(* IEC 61131-3 sources: PortalRobot/Portal_robot/Device/application/ST/ST_CELL, 17 files *)

(* ---- E_CELL_MANAGER_STATE.st ---- *)
{attribute 'qualified_only'}
{attribute 'strict'}
TYPE E_CELL_MANAGER_STATE :
(
	IDLE,
	PLAN_TARGET,
	MAGAZINE_EXECUTE,
	RELEASE_MAGAZINE,
	ROUTE_TO_TARGET,
	RELEASE_ROBOT_COMMAND,
	WAIT_TARGET,
	SERVICE_TARGET,
	SELECT_FALLBACK,
	WAIT_MAGAZINE,
	ERROR,
	MACHINE_FAULT_STOP,
	PRESTART_IDENTIFY,
	WAIT_GRIPPER1_CONTENT,
	WAIT_GRIPPER1_TYPE,
	WAIT_GRIPPER2_CONTENT,
	WAIT_GRIPPER2_TYPE,
	WAIT_START_MACHINE,
	TEST_ABORT_STOP,
	GEOMETRY_WAIT_FREE,
	GEOMETRY_DELIVER,
	GEOMETRY_RELEASE_COMMAND
);
END_TYPE

(* ---- E_CELL_STATE.st ---- *)
{attribute 'qualified_only'}
{attribute 'strict'}
TYPE E_CELL_STATE :
(
	IDLE,
	ROUTE_PAYLOAD,
	SELECT_MACHINE,
	MOVE_TO_MACHINE,
	RELEASE_ROBOT_COMMAND,
	WAIT_MACHINE,
	SERVICE_MACHINE,
	MAGAZINE,
	RELEASE_MAGAZINE,
	WAIT_MAGAZINE,
	ERROR,
	GEOMETRY_WAIT,
	GEOMETRY_TRANSFER
);
END_TYPE

(* ---- ST_BUTTON_STATION_IO_STATUS.st ---- *)
TYPE ST_BUTTON_STATION_IO_STATUS :
STRUCT
	xEmergencyStopPressed : BOOL; // Нормализованный вход: TRUE — грибок нажат
	xButtonPressed        : BOOL; // Нормализованный вход кнопки открытия замка
	xButtonLightOn        : BOOL; // Фактический выход подсветки кнопки
END_STRUCT
END_TYPE

(* ---- ST_CELL_COMMAND.st ---- *)
TYPE ST_CELL_COMMAND :
STRUCT
	stRobot          : ST_ROBOT_COMMAND; // Команда роботу от менеджера ячейки
	uiBlankPayloadType  : UINT; // Тип заготовки в первом захвате
	uiDetailPayloadType : UINT; // Тип готовой детали во втором захвате
	stMagazine       : ST_MAGAZINE_COMMAND; // Команда магазину
	axMachineExecute : ARRAY [1..3] OF BOOL; // Запуск обслуживания выбранного станка
END_STRUCT
END_TYPE

(* ---- ST_CELL_CYCLE_STATUS.st ---- *)
TYPE ST_CELL_CYCLE_STATUS :
STRUCT
	eState              : E_CELL_MANAGER_STATE; // Состояние универсального автомата ячейки
	uiSelectedMachine   : UINT; // Зафиксированный целевой станок
	uiSelectedType      : UINT; // Тип заготовки текущего маршрута
	uiBlankPayloadType  : UINT; // Тип заготовки в первом захвате
	uiDetailPayloadType : UINT; // Тип готовой детали во втором захвате
	iTakeSlot           : SINT; // Зарезервированный слот взятия
	iPutSlot            : SINT; // Зарезервированный слот укладки
	xReturningBlank     : BOOL; // Выполняется возврат заготовки
	axMachineStartPending: ARRAY [1..3] OF BOOL; // Запуск нового цикла ещё подтверждается станком
	auiBlankCount       : ARRAY [1..3] OF UINT; // Заготовки по типам
	auiDetailCount      : ARRAY [1..3] OF UINT; // Готовые детали по типам
	auiFreeCount        : ARRAY [1..3] OF UINT; // Свободные слоты по типам
END_STRUCT
END_TYPE

(* ---- ST_CELL_DIAG.st ---- *)
TYPE ST_CELL_DIAG :
STRUCT
	eState : E_CELL_STATE; // Текущее состояние автомата ячейки
	stWarning : ST_WARNING_EVENT; // Последнее предупреждение менеджера ячейки
END_STRUCT
END_TYPE

(* ---- ST_CELL_ERROR.st ---- *)
TYPE ST_CELL_ERROR :
STRUCT
	BOTH_GRIPPERS_OCCUPIED : BOOL; // Совместимый бит: диагностическая ошибка согласованности захватов
	ROBOT_ERROR            : BOOL; // Ошибка робота во время автоматического цикла
	MAGAZINE_ERROR         : BOOL; // Ошибка магазина во время операции
	MACHINE_ERROR          : BOOL; // Ошибка станка во время обслуживания
	GLOBAL_STOP            : BOOL; // Получена глобальная ошибка ячейки
END_STRUCT
END_TYPE

(* ---- ST_CELL_ERRORS.st ---- *)
TYPE ST_CELL_ERRORS :
STRUCT
	dwErrorActive : DWORD; // Битовая маска активных ошибок
	dwErrorLast   : DWORD; // Битовая маска последних ошибок
	dwAlarmActive : DWORD; // Собственные аварии менеджера ячейки для общего журнала
	stErrorActive : ST_CELL_ERROR; // Расшифровка активных ошибок
	stErrorLast   : ST_CELL_ERROR; // Расшифровка последних ошибок
END_STRUCT
END_TYPE

(* ---- ST_CELL_FAULT_REQUEST.st ---- *)
TYPE ST_CELL_FAULT_REQUEST :
STRUCT
	xEnabled      : BOOL; // Глобальное разрешение диагностической инъекции
	xBothGrippers : BOOL; // Совместимый диагностический импульс ошибки согласованности захватов
END_STRUCT
END_TYPE

(* ---- ST_CELL_SAFETY_DIAG.st ---- *)
TYPE ST_CELL_SAFETY_DIAG :
STRUCT
	stWarning : ST_WARNING_EVENT; // Отклонённые попытки открытия и сброса реле
END_STRUCT
END_TYPE

(* ---- ST_CELL_SAFETY_ERRORS.st ---- *)
TYPE ST_CELL_SAFETY_ERRORS :
STRUCT
	dwErrorActive : DWORD; // Текущие отдельные Safety-причины
	dwErrorLast   : DWORD; // Последняя ненулевая маска для диагностики
	dwAlarmActive : DWORD; // Собственные аварии источника для общего журнала
END_STRUCT
END_TYPE

(* ---- ST_CELL_SAFETY_FAULT_REQUEST.st ---- *)
TYPE ST_CELL_SAFETY_FAULT_REQUEST :
STRUCT
	xEnabled : BOOL; // Общее разрешение диагностических инъекций
	axEmergencyStopStation : ARRAY [1..4] OF BOOL;
	axEmergencyStopCabinet : ARRAY [1..2] OF BOOL;
	xEmergencyStopMpg      : BOOL;
	xPhaseRelayFault       : BOOL;
	xPressureRelayFault    : BOOL;
	xSafetyRelayFault      : BOOL;
	axDoorUnlocked         : ARRAY [1..4] OF BOOL;
END_STRUCT
END_TYPE

(* ---- ST_CELL_SAFETY_STATUS.st ---- *)
TYPE ST_CELL_SAFETY_STATUS :
STRUCT
	xReady                   : BOOL; // Все текущие условия безопасности выполнены
	xGlobalError             : BOOL; // Хотя бы одна текущая Safety-причина активна
	xPhaseRelayOk            : BOOL; // Реле контроля фаз в норме
	xPressureRelayOk         : BOOL; // Реле контроля давления в норме
	xSafetyRelayOk           : BOOL; // Реле безопасности взведено
	xSafetyRelayResetAllowed : BOOL; // Разрешён отдельный импульс сброса реле
	xSafetyRelayResetActive  : BOOL; // Полный секундный импульс сброса реле сейчас активен
	axEmergencyStopReleased  : ARRAY [1..7] OF BOOL; // 4 поста, 2 шкафа, MPG
	axDoorReady              : ARRAY [1..4] OF BOOL; // Замок закрыт либо связанный магазин выключен
	axButtonStationPressed   : ARRAY [1..4] OF BOOL; // Фактический вход кнопки поста, с учётом симуляции
	axButtonStationLightOn   : ARRAY [1..4] OF BOOL; // Выход подсветки кнопки поста
END_STRUCT
END_TYPE

(* ---- ST_CELL_STATUS.st ---- *)
TYPE ST_CELL_STATUS :
STRUCT
	xMagazineExchangeAllowed : BOOL; // Планировщик не держит незавершённый маршрут
	xRunning           : BOOL; // Автоматический цикл запущен
	xStopPending       : BOOL; // Запрошена остановка после безопасного шага
	xBusy              : BOOL; // Менеджер выполняет автоматический цикл
	xWaitingMachine    : BOOL; // Ожидание доступного станка
	xWaitingMagazine   : BOOL; // Ожидание пополнения или освобождения магазина
	xError             : BOOL; // Менеджер ячейки находится в ошибке
	xReadyToStart      : BOOL; // Выполнены все условия запуска автоматического цикла
	xStartAllowed      : BOOL; // Кнопка запуска или отмены ожидающей остановки доступна
	xStopAllowed       : BOOL; // Кнопка остановки автоматического цикла доступна
	xResetAllowed      : BOOL; // Кнопка общего сброса доступна
	xManualAllowed     : BOOL; // Кнопка перехода в ручной режим доступна
	xAutomaticAllowed  : BOOL; // Кнопка перехода в автоматический режим доступна
	xDrivesReady       : BOOL; // Приводы и группа осей готовы к движению
	xRobotReady        : BOOL; // Робот готов принять команду
	xMagazineReady     : BOOL; // Магазин готов к работе с роботом
	xSafetyHomeRequired: BOOL; // Повторный запуск разрешён только из HOME_SAFETY
	xRobotAtSafetyHome : BOOL; // Фактические координаты находятся в диапазоне HOME_SAFETY
	xStartCheckCellIdle          : BOOL; // Менеджер ячейки готов принять новый запуск
	xStartCheckAutomaticMode     : BOOL; // Выбран автоматический режим
	xStartCheckNoBlockingError   : BOOL; // Нет блокирующей запуск ошибки
	xStartCheckRobotInterfaceReady: BOOL; // Выбранный интерфейс робота готов
	xStartCheckConfigurationValid: BOOL; // Конфигурация типов корректна
	xStartCheckPointsConfigured  : BOOL; // HOME_SAFETY и точки включённого оборудования настроены
	xStartCheckDrivesReady       : BOOL; // Приводы и группа готовы
	xStartCheckRobotReady        : BOOL; // Робот готов принять маршрут
	xStartCheckMagazineReady     : BOOL; // Магазин готов к операции
	xStartCheckTaskAvailable     : BOOL; // Есть допустимая работа или известный груз
	xStartCheckSafetyHome        : BOOL; // Условие HOME_SAFETY выполнено
	xStartCheckSafety            : BOOL; // Грибки, реле и двери безопасности готовы
	uiStartConditionsMet        : UINT; // Количество выполненных условий запуска
	uiStartConditionsTotal      : UINT; // Общее количество условий запуска
	uiReadyMachines    : UINT; // Количество включённых станков в состоянии IDLE
	uiSelectedMachine  : UINT; // Номер выбранного станка
	uiActiveMagazine   : UINT; // Магазин, закреплённый за текущим автоматическим циклом
	eMagazineOperation : E_MAGAZINE_OPERATION; // Выбранная операция магазина
	xOperatorPromptActive : BOOL; // PLC ожидает ответ оператора перед запуском цикла
	xOperatorChoiceAllowed: BOOL; // PLC разрешает отправить вариант активного опроса
	xOperatorCancelAllowed: BOOL; // PLC разрешает отменить активный предпусковой опрос
	uiOperatorPrompt      : UINT; // 0 нет; 1/3 содержимое захвата; 2/4 тип; 5 станок
	uiOperatorTypeMask    : UINT; // Биты 0..2 — доступные типы продукции
	uiOperatorMachineMask : UINT; // Биты 0..2 — допустимые станки для стартового LOAD
END_STRUCT
END_TYPE

(* ---- ST_CONTROL_CABINET_IO_STATUS.st ---- *)
TYPE ST_CONTROL_CABINET_IO_STATUS :
STRUCT
	xEmergencyStopPressed : BOOL; // Нормализованный вход: TRUE — грибок нажат
	xStartPressed         : BOOL; // Физическая кнопка «Включить ячейку»
	xStopPressed          : BOOL; // Физическая кнопка «Выключить ячейку»
	xResetPressed         : BOOL; // Физическая кнопка общего сброса ошибок
END_STRUCT
END_TYPE

(* ---- ST_ENCLOSURE_DOOR_STATUS.st ---- *)
TYPE ST_ENCLOSURE_DOOR_STATUS :
STRUCT
	xLocked        : BOOL; // Обратная связь замка: TRUE — замок закрыт
	xUnlockAllowed : BOOL; // PLC разрешает открыть замок
	xUnlockOutput  : BOOL; // Фактическая команда открытия замка
END_STRUCT
END_TYPE

(* ---- ST_MPG_IO_STATUS.st ---- *)
TYPE ST_MPG_IO_STATUS :
STRUCT
	xEmergencyStopPressed : BOOL; // Нормализованный вход: TRUE — грибок MPG нажат
	xAxisX                : BOOL; // Положение селектора оси X
	xAxisY                : BOOL; // Положение селектора оси Y
	xAxisZ                : BOOL; // Положение селектора оси Z
	xMultiplier1          : BOOL; // Положение множителя x1
	xMultiplier10         : BOOL; // Положение множителя x10
	xMultiplier100        : BOOL; // Положение множителя x100
END_STRUCT
END_TYPE
